(* Schneider Machine Expert - Basic project register_fifo_m20_m21_m22_contacts_il_only, file version 3.0.0.0 *)
(* ProjectInformations: Name=New project *)

HARDWARE
  Cpu 0: TM200CE40T
  EthernetConfiguration: NetworkName=M200, IpAllocationMode=FixedAddress, IpAddress=0.0.0.0, SubnetMask=0.0.0.0
  SerialLineConfiguration: Baud=Baud19200, Parity=ParityEven, DataBits=DataBits8, StopBits=StopBits1, PhysicalMedium=PhysicalMediumRs485, TransmissionMode=TransmissionModeModbusRtu, SlaveId=1, Addressing=SlaveAddressing
  MastTask: UsePeriodScanMode=false, PeriodScan=100
  FastTask: Period=255
  CpuBehavior: StartingMode=StartAsPreviousState, AutoSaveRamOnEeprom=true, WatchdogPeriod=250

SYMBOLS  (address, symbol, comment, settings)

POU New POU
  (* SectionNumber=0 *)

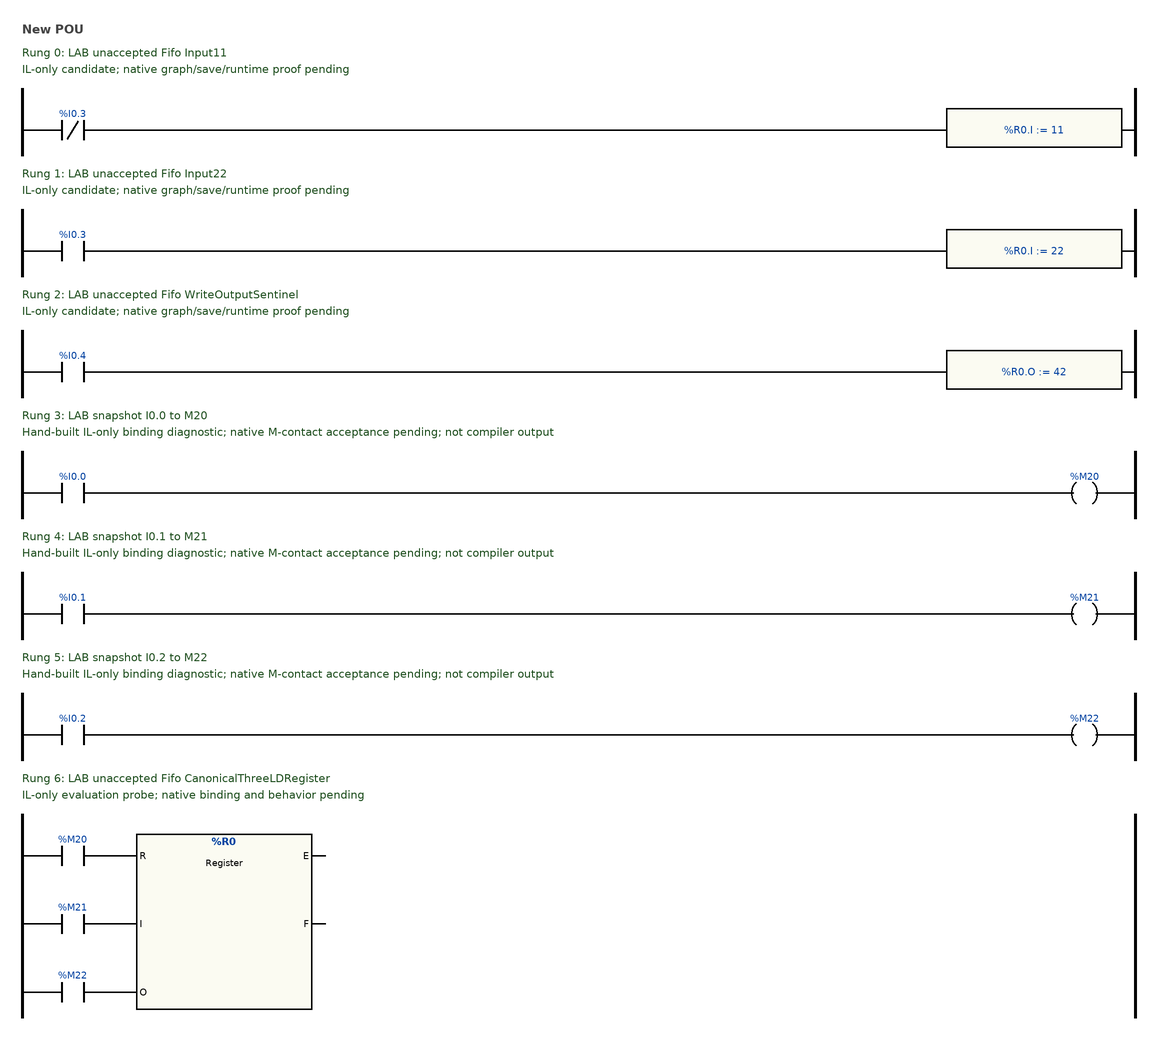

// Rung 0: LAB unaccepted Fifo Input11
// IL-only candidate; native graph/save/runtime proof pending
  LDN %I0.3
  [ %R0.I := 11 ]
  // as ST:
  //   IF NOT %I0.3 THEN %R0.I := 11; END_IF;

// Rung 1: LAB unaccepted Fifo Input22
// IL-only candidate; native graph/save/runtime proof pending
  LD %I0.3
  [ %R0.I := 22 ]
  // as ST:
  //   IF %I0.3 THEN %R0.I := 22; END_IF;

// Rung 2: LAB unaccepted Fifo WriteOutputSentinel
// IL-only candidate; native graph/save/runtime proof pending
  LD %I0.4
  [ %R0.O := 42 ]
  // as ST:
  //   IF %I0.4 THEN %R0.O := 42; END_IF;

// Rung 3: LAB snapshot I0.0 to M20
// Hand-built IL-only binding diagnostic; native M-contact acceptance pending; not compiler output
  LD %I0.0
  ST %M20
  // as ST:
  //   %M20 := %I0.0;

// Rung 4: LAB snapshot I0.1 to M21
// Hand-built IL-only binding diagnostic; native M-contact acceptance pending; not compiler output
  LD %I0.1
  ST %M21
  // as ST:
  //   %M21 := %I0.1;

// Rung 5: LAB snapshot I0.2 to M22
// Hand-built IL-only binding diagnostic; native M-contact acceptance pending; not compiler output
  LD %I0.2
  ST %M22
  // as ST:
  //   %M22 := %I0.2;

// Rung 6: LAB unaccepted Fifo CanonicalThreeLDRegister
// IL-only evaluation probe; native binding and behavior pending
  BLK %R0
  LD %M20
  R
  LD %M21
  I
  LD %M22
  O
  END_BLK
  // as ST:
  //   %R0(R := %M20, I := %M21, O := %M22);

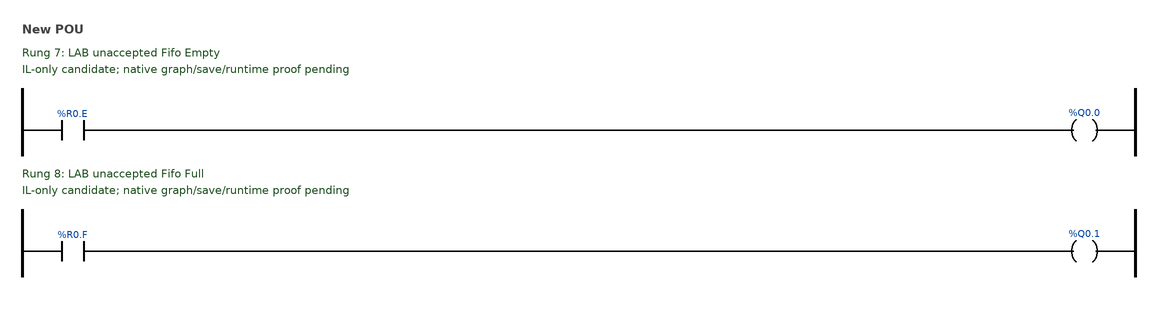

// Rung 7: LAB unaccepted Fifo Empty
// IL-only candidate; native graph/save/runtime proof pending
  LD %R0.E
  ST %Q0.0
  // as ST:
  //   %Q0.0 := %R0.E;

// Rung 8: LAB unaccepted Fifo Full
// IL-only candidate; native graph/save/runtime proof pending
  LD %R0.F
  ST %Q0.1
  // as ST:
  //   %Q0.1 := %R0.F;
